(* PLC project PR_5by3CylModWoRdlck_PLC, SiemensToBackhoff Siemens TIA Portal to Beckhoff TwinCAT PLCopen Converter 2.0 *)
(* stored: creationDateTime 2026-09-28T12:19:39.070834, modificationDateTime 2026-09-28T12:19:39.070834 *)

FUNCTION_BLOCK PR_5by3CylModWoRdlck
VAR_INPUT
	iResetModule : BOOL;  // Reset if 1
	iResetFaults : BOOL;  // Reset Fault CMD
	iEnergizeAtPwrOn : BOOL;  // Energize Poweron Input
	iWorkCmd : BOOL;  // Cyl Work Postion CMD
	iHomeCmd : BOOL;  // Cyl Home Postion CMD
	iWorkSen : BOOL;  // Cyl Work Postion Input
	iHomeSen : BOOL;  // Cyl Home Postion Input
	iWorkCleartoMove : BOOL;  // connect work position interlock condition healthy
	iHomeCleartoMove : BOOL;  // connect home position interlock condition healthy
	iWorkPositionLeftOption : BOOL;  // It is the selection of the to keep work solenoid coil on after reaching work position
	iHomePositionLeftOption : BOOL;  // It is the selection of the to keep home solenoid coil on after reaching home position
	iTimeoutValue : TIME;  // Time Required E.g T#500MS,T#2S
	iWorkSensDebounceVal : TIME;  // Time Required E.g T#500MS,T#2S
	iHomeSensDebounceVal : TIME;  // Time Required E.g T#500MS,T#2S
END_VAR
VAR_OUTPUT
	qWorkSol : BOOL;  // Cyl Work Position Sol Output
	qHomeSol : BOOL;  // Cyl Home Position Sol Output
	qWorkOver : BOOL;  // 1 if Cyl at Work Position
	qHomeOver : BOOL;  // 1 if Cyl at Home Position
	qModError : BOOL;  // Module Error
	qErrBothSensorOn : BOOL;  // 1 If both WorkSen and HomeSen inputs are high at the same time.
	qErrHomeInterlock : BOOL;  // 1 If homeCleartoMove is low and home command is active.
	qErrHomeSenNotLeft : BOOL;  // 1 If home position sensor did not turn off within defined time
	qErrHomeTout : BOOL;  // 1 If cylinder did not reach home position within defined time
	qErrWorkInterlock : BOOL;  // 1 If WorkCleartoMove is low and work command is active.
	qErrWorkSenNotLeft : BOOL;  // 1 If work position sensor did not turn off within defined time
	qErrWorkTout : BOOL;  // 1 If cylinder did not reach work position within defined time
	qMsgWorkPosLost : BOOL;  // 1 If work position achieved and lost its position without home
	qMsgHomePosLost : BOOL;  // 1 If home position achieved and lost its position without work
	qMsgBothCmdOn : BOOL;  // 1 if Home & work position command on same time
END_VAR
VAR
	sFltRstPls : BOOL;  // Stat bit for positive edge of reset fault input
	sFltEdge : R_TRIG;  // Positive edge of fault reset input
	sWorkPosMemBit : BOOL;  // Stat bit for work position memory bit
	sHomePosMemBit : BOOL;  // Stat bit for Home position memory bit
	sModError : BOOL;  // Stat bit for Module error
	sWorkSensDebTime : TIME;  // Stat bit work sensor debounce time
	sHomeSensDebTime : TIME;  // Stat bit work sensor debounce time
	sTimeoutValue : TIME;  // Stat bit for time out value
	sElapsedTime : TIME;  // Stat bit for time elapsed
	sDlyWorkSensDeb : TON;  // On Delay for Work Sensor Debounce
	sDlyHomeSensDeb : TON;  // On Delay For Home Sensor Debounce
	sDlyTimeOut : TON;  // On Delay Time Out timer
	sWorkSol : BOOL;
	sErrWorkTout : BOOL;
	sHomeSol : BOOL;
	sErrHomeTout : BOOL;
	sErrBothSensorOn : BOOL;
	sErrWorkInterlock : BOOL;
	sErrHomeInterlock : BOOL;
	sErrWorkSenNotLeft : BOOL;
	sErrHomeSenNotLeft : BOOL;
	sMsgHomePosLost : BOOL;
	sMsgWorkPosLost : BOOL;
	sPosEdge : R_TRIG;
	sPosEdge1 : R_TRIG;
	sRegainWrkPos : BOOL;
	sRegainHomePos : BOOL;
	sBothCmdOn : BOOL;
	sWorkPositionLeft : BOOL;
	sHomePositionLeft : BOOL;
END_VAR
  VAR  (* added by the conversion: wires and edge detectors of the diagram *)
    _EQ31_ENO : BOOL;
    _EQ31_OUT : BOOL;
    _EQ47_ENO : BOOL;
    _EQ47_OUT : BOOL;
    _EQ63_ENO : BOOL;
    _EQ63_OUT : BOOL;
  END_VAR

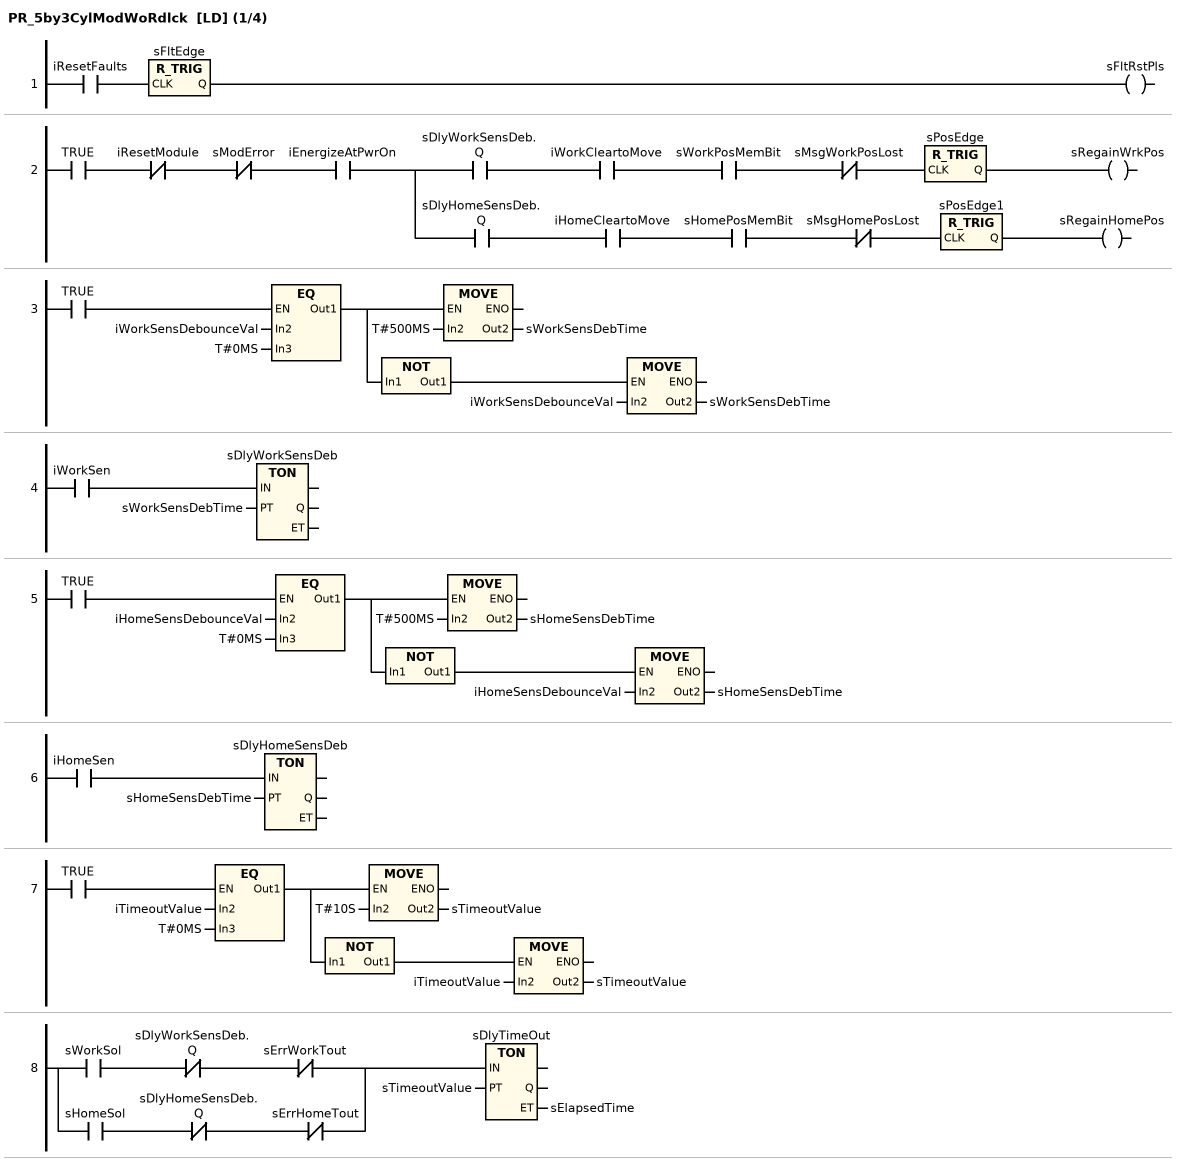
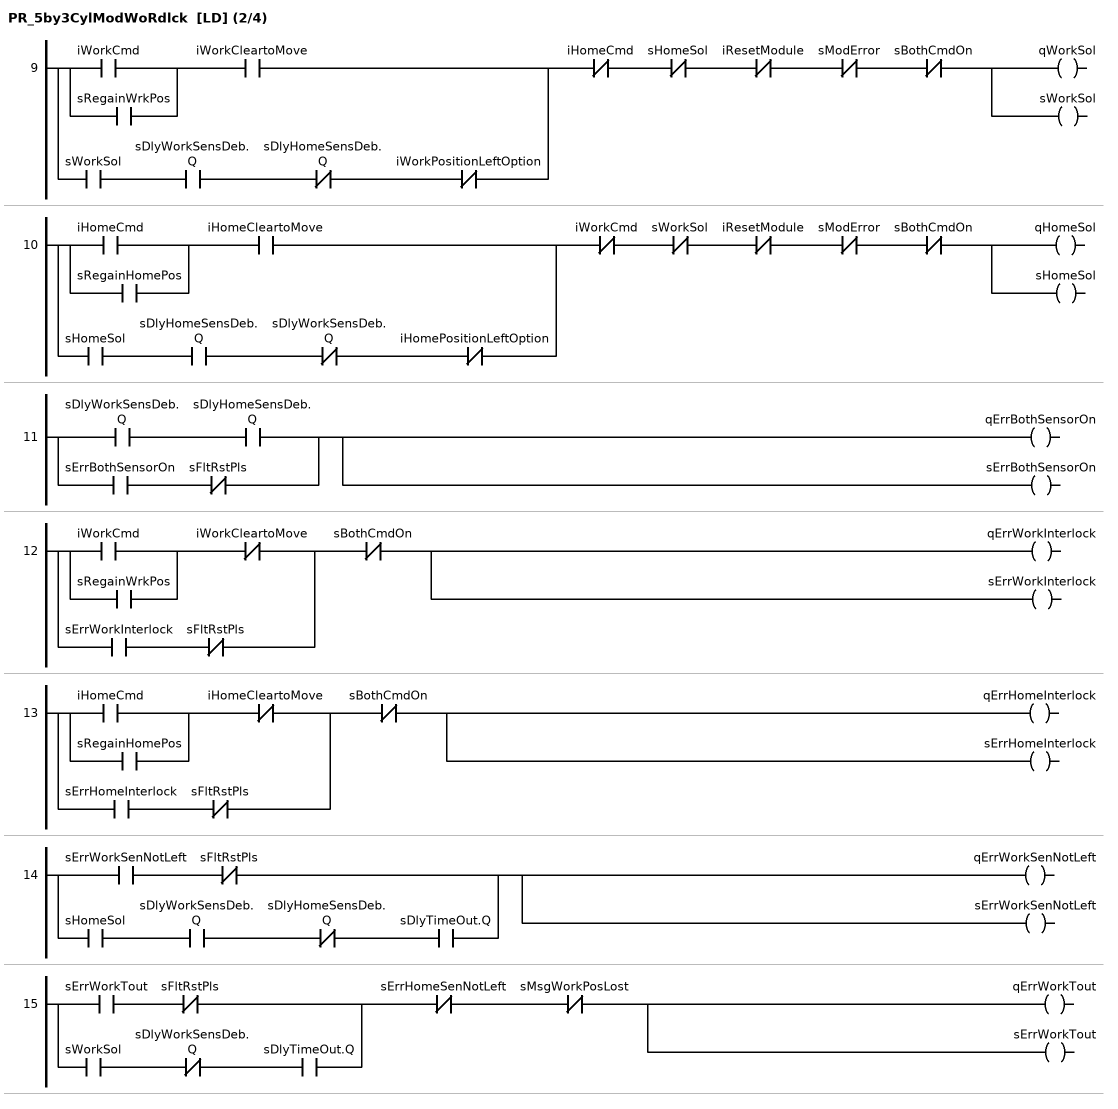
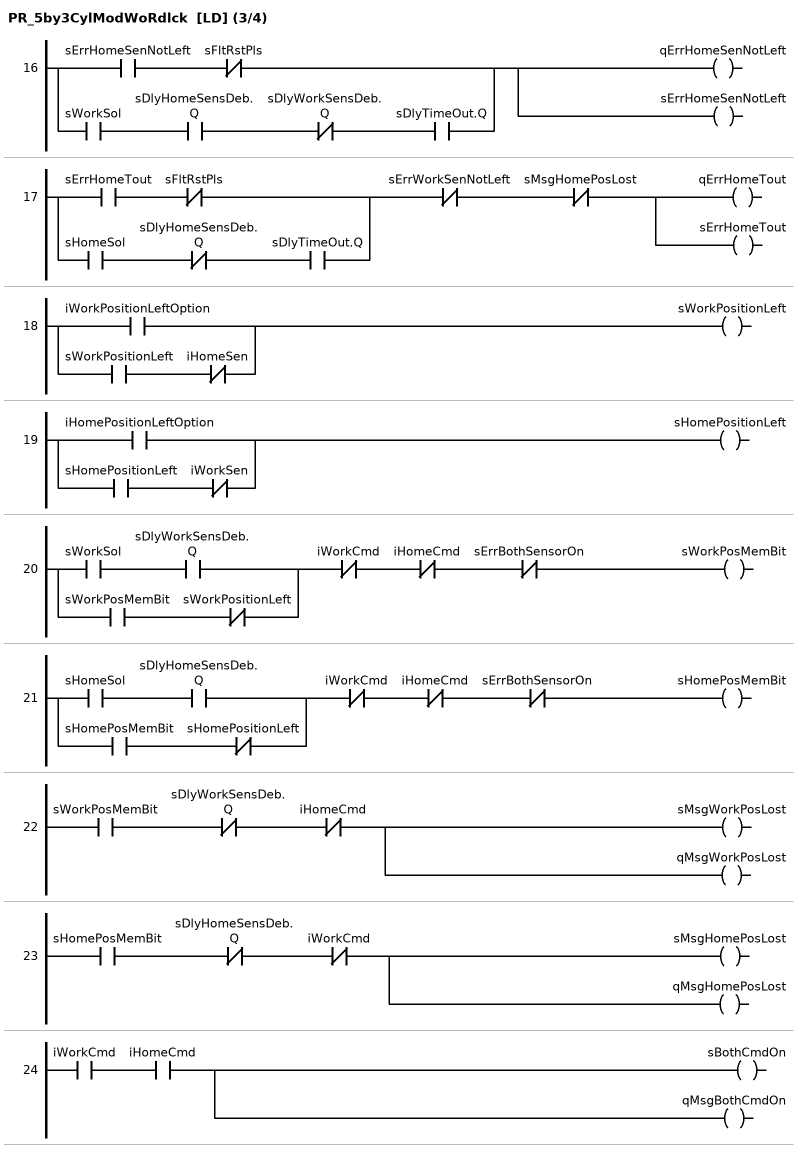
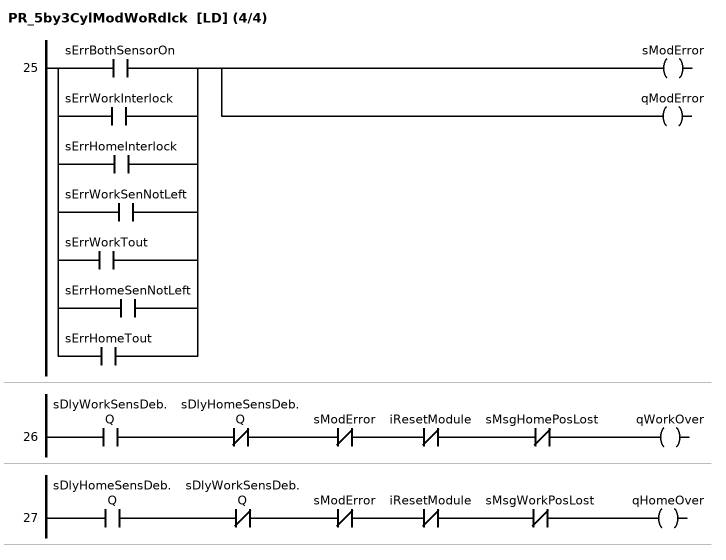
(* LD diagram, written out as Structured Text *)
(* ==============================================================================
 Company: Precision Automation & Robotics India Ltd. 
------------------------------------------------------------------------------
 Item Code:SM0101022005
 Author/Created by: Amiya Das
 Reviewed/Checked by: Atul Patwardhan
 First Release on: 20-01-2017
 Latest update on:27-01-2025 
------------------------------------------------------------------------------
 Tested with:Simulator
 Engineering/Editor: TIA Portal 15 & Higher
------------------------------------------------------------------------------
 Restrictions: No
 Dependencies/Requirements: NA
------------------------------------------------------------------------------
 Change Log:
 Ver.	Date                            Changed by                                  Details of changes
 0.2           20-01-2017                  Amiya Das      	              Second release version
 0.3           27-01-2025                 Sujeet Rote                                qMsgBothCmdOn message is added
 0.4           29-01-2025                  Sujeet Rote                                Work & home position left option bit
------------------------------------------------------------------------------
Functionality: This block is used to control a simple motion with one work 
position output, one home position  output, one work position sensor and one 
home position sensor.
Inputs
iResetModule	Bool
iResetFaults	Bool
iEnergizeAtPwrOn	Bool
iWorkCmd	Bool
iHomeCmd	Bool
iWorkSen	Bool
iHomeSen	Bool
iWorkCleartoMove	Bool
iHomeCleartoMove	Bool
iWorkPositionLeftOption	Bool
iHomePositionLeftOption	Bool
iTimeoutValue	Time
iWorkSensDebounceVal	Time
iHomeSensDebounceVal	Time

Outputs
qWorkSol	Bool
qHomeSol	Bool
qWorkOver	Bool
qHomeOver	Bool
qErrBothSensorOn	Bool
qErrHomeInterlock	Bool
qErrHomeSenNotLeft	Bool
qErrHomeTout	Bool
qErrWorkInterlock	Bool
qErrWorkSenNotLeft	Bool
qErrWorkTout	Bool
qMsgWorkPosLost	Bool
qMsgHomePosLost	Bool
qMsgBothCmdOn	Bool

In-outs
NIL
------------------------------------------------------------------------------
Errors reported:
1.qErrBothSensorOn: If both WorkSen and HomeSen inputs are high at the same time.          
2.qErrHomeInterlock: If homeCleartoMove is low and home command is active.
3.qErrHomeSenNotLeft: If home position sensor did not turn off within defined time 
4.qErrHomeTout: If cylinder did not reach home position within defined time 
5.qErrWorkInterlock: If WorkCleartoMove is low and work command is active. 
7.qErrWorkSenNotLeft: If work position sensor did not turn off within defined time 
8.qErrWorkTout: If cylinder did not reach work position within defined time 
9.qErrPipeSwaped: If Pipe or sensor swapped

Messages reported:
1.qMsgHomePosLost: If home position achieved and lost its position without work
2.qMsgWorkPosLost: If work position achieved and lost its position without home 
3.qMsgBothCmdOn :  Home & work position command on same time
============================================================================== *)

(* Fault Reset Pulse *)

sFltEdge(CLK := iResetFaults);
sFltRstPls := sFltEdge.Q;
(* Regain Position after power On logic *)

sPosEdge(CLK := TRUE AND NOT iResetModule AND NOT sModError AND iEnergizeAtPwrOn AND sDlyWorkSensDeb.Q AND iWorkCleartoMove AND sWorkPosMemBit AND NOT sMsgWorkPosLost);
sRegainWrkPos := sPosEdge.Q;
sPosEdge1(CLK := TRUE AND NOT iResetModule AND NOT sModError AND iEnergizeAtPwrOn AND sDlyHomeSensDeb.Q AND iHomeCleartoMove AND sHomePosMemBit AND NOT sMsgHomePosLost);
sRegainHomePos := sPosEdge1.Q;
(* Work sensor default debounce value *)

_EQ31_OUT := EQ(EN := TRUE, IN1 := iWorkSensDebounceVal, IN2 := T#0MS, ENO => _EQ31_ENO);
IF _EQ31_OUT THEN sWorkSensDebTime := T#500MS; END_IF;
IF NOT _EQ31_OUT THEN sWorkSensDebTime := iWorkSensDebounceVal; END_IF;
(* Work Sensor On Debounce Timer *)

sDlyWorkSensDeb(IN := iWorkSen, PT := sWorkSensDebTime);
(* Home sensor default debounce value *)

_EQ47_OUT := EQ(EN := TRUE, IN1 := iHomeSensDebounceVal, IN2 := T#0MS, ENO => _EQ47_ENO);
IF _EQ47_OUT THEN sHomeSensDebTime := T#500MS; END_IF;
IF NOT _EQ47_OUT THEN sHomeSensDebTime := iHomeSensDebounceVal; END_IF;
(* Home Sensor On Debounce Timer *)

sDlyHomeSensDeb(IN := iHomeSen, PT := sHomeSensDebTime);
(* Timeout Value *)

_EQ63_OUT := EQ(EN := TRUE, IN1 := iTimeoutValue, IN2 := T#0MS, ENO => _EQ63_ENO);
IF _EQ63_OUT THEN sTimeoutValue := T#10S; END_IF;
IF NOT _EQ63_OUT THEN sTimeoutValue := iTimeoutValue; END_IF;
(* Sensor timeout Timer *)

sDlyTimeOut(IN := sWorkSol AND NOT sDlyWorkSensDeb.Q AND NOT sErrWorkTout OR sHomeSol AND NOT sDlyHomeSensDeb.Q AND NOT sErrHomeTout, PT := sTimeoutValue, ET => sElapsedTime);
(* Cylinder Work Sol *)

qWorkSol := ((iWorkCmd OR sRegainWrkPos) AND iWorkCleartoMove OR sWorkSol AND sDlyWorkSensDeb.Q AND NOT sDlyHomeSensDeb.Q AND NOT iWorkPositionLeftOption) AND NOT iHomeCmd AND NOT sHomeSol AND NOT iResetModule AND NOT sModError AND NOT sBothCmdOn;
sWorkSol := ((iWorkCmd OR sRegainWrkPos) AND iWorkCleartoMove OR sWorkSol AND sDlyWorkSensDeb.Q AND NOT sDlyHomeSensDeb.Q AND NOT iWorkPositionLeftOption) AND NOT iHomeCmd AND NOT sHomeSol AND NOT iResetModule AND NOT sModError AND NOT sBothCmdOn;
(* Cylinder Home Sol *)

qHomeSol := ((iHomeCmd OR sRegainHomePos) AND iHomeCleartoMove OR sHomeSol AND sDlyHomeSensDeb.Q AND NOT sDlyWorkSensDeb.Q AND NOT iHomePositionLeftOption) AND NOT iWorkCmd AND NOT sWorkSol AND NOT iResetModule AND NOT sModError AND NOT sBothCmdOn;
sHomeSol := ((iHomeCmd OR sRegainHomePos) AND iHomeCleartoMove OR sHomeSol AND sDlyHomeSensDeb.Q AND NOT sDlyWorkSensDeb.Q AND NOT iHomePositionLeftOption) AND NOT iWorkCmd AND NOT sWorkSol AND NOT iResetModule AND NOT sModError AND NOT sBothCmdOn;
(* Both Sensor On Error *)

qErrBothSensorOn := sDlyWorkSensDeb.Q AND sDlyHomeSensDeb.Q OR sErrBothSensorOn AND NOT sFltRstPls;
sErrBothSensorOn := sDlyWorkSensDeb.Q AND sDlyHomeSensDeb.Q OR sErrBothSensorOn AND NOT sFltRstPls;
(* Work Interlock Error *)

qErrWorkInterlock := ((iWorkCmd OR sRegainWrkPos) AND NOT iWorkCleartoMove OR sErrWorkInterlock AND NOT sFltRstPls) AND NOT sBothCmdOn;
sErrWorkInterlock := ((iWorkCmd OR sRegainWrkPos) AND NOT iWorkCleartoMove OR sErrWorkInterlock AND NOT sFltRstPls) AND NOT sBothCmdOn;
(* Home Interlock Error pending *)

qErrHomeInterlock := ((iHomeCmd OR sRegainHomePos) AND NOT iHomeCleartoMove OR sErrHomeInterlock AND NOT sFltRstPls) AND NOT sBothCmdOn;
sErrHomeInterlock := ((iHomeCmd OR sRegainHomePos) AND NOT iHomeCleartoMove OR sErrHomeInterlock AND NOT sFltRstPls) AND NOT sBothCmdOn;
(* Work Sensor Not Left Error  pending *)

qErrWorkSenNotLeft := sHomeSol AND sDlyWorkSensDeb.Q AND NOT sDlyHomeSensDeb.Q AND sDlyTimeOut.Q OR sErrWorkSenNotLeft AND NOT sFltRstPls;
sErrWorkSenNotLeft := sHomeSol AND sDlyWorkSensDeb.Q AND NOT sDlyHomeSensDeb.Q AND sDlyTimeOut.Q OR sErrWorkSenNotLeft AND NOT sFltRstPls;
(* Work Timeout Error *)

qErrWorkTout := (sWorkSol AND NOT sDlyWorkSensDeb.Q AND sDlyTimeOut.Q OR sErrWorkTout AND NOT sFltRstPls) AND NOT sErrHomeSenNotLeft AND NOT sMsgWorkPosLost;
sErrWorkTout := (sWorkSol AND NOT sDlyWorkSensDeb.Q AND sDlyTimeOut.Q OR sErrWorkTout AND NOT sFltRstPls) AND NOT sErrHomeSenNotLeft AND NOT sMsgWorkPosLost;
(* Home Sensor Not Left Error *)

qErrHomeSenNotLeft := sWorkSol AND sDlyHomeSensDeb.Q AND NOT sDlyWorkSensDeb.Q AND sDlyTimeOut.Q OR sErrHomeSenNotLeft AND NOT sFltRstPls;
sErrHomeSenNotLeft := sWorkSol AND sDlyHomeSensDeb.Q AND NOT sDlyWorkSensDeb.Q AND sDlyTimeOut.Q OR sErrHomeSenNotLeft AND NOT sFltRstPls;
(* Home Timeout Error *)

qErrHomeTout := (sHomeSol AND NOT sDlyHomeSensDeb.Q AND sDlyTimeOut.Q OR sErrHomeTout AND NOT sFltRstPls) AND NOT sErrWorkSenNotLeft AND NOT sMsgHomePosLost;
sErrHomeTout := (sHomeSol AND NOT sDlyHomeSensDeb.Q AND sDlyTimeOut.Q OR sErrHomeTout AND NOT sFltRstPls) AND NOT sErrWorkSenNotLeft AND NOT sMsgHomePosLost;
(* Work Position Left option bit Logic *)

sWorkPositionLeft := iWorkPositionLeftOption OR sWorkPositionLeft AND NOT iHomeSen;
(* Home Position Left option bit Logic *)

sHomePositionLeft := iHomePositionLeftOption OR sHomePositionLeft AND NOT iWorkSen;
(* Work Position Memory Bit *)

sWorkPosMemBit := (sWorkSol AND sDlyWorkSensDeb.Q OR sWorkPosMemBit AND NOT sWorkPositionLeft) AND NOT iWorkCmd AND NOT iHomeCmd AND NOT sErrBothSensorOn;
(* Home Position Memory Bit *)

sHomePosMemBit := (sHomeSol AND sDlyHomeSensDeb.Q OR sHomePosMemBit AND NOT sHomePositionLeft) AND NOT iWorkCmd AND NOT iHomeCmd AND NOT sErrBothSensorOn;
(* Msg:-Work Position Lost *)

sMsgWorkPosLost := sWorkPosMemBit AND NOT sDlyWorkSensDeb.Q AND NOT iHomeCmd;
qMsgWorkPosLost := sWorkPosMemBit AND NOT sDlyWorkSensDeb.Q AND NOT iHomeCmd;
(* Msg:- Home Position Lost *)

sMsgHomePosLost := sHomePosMemBit AND NOT sDlyHomeSensDeb.Q AND NOT iWorkCmd;
qMsgHomePosLost := sHomePosMemBit AND NOT sDlyHomeSensDeb.Q AND NOT iWorkCmd;
(* Msg:- Both command On *)

sBothCmdOn := iWorkCmd AND iHomeCmd;
qMsgBothCmdOn := iWorkCmd AND iHomeCmd;
(* Module Error *)

sModError := sErrBothSensorOn OR sErrWorkInterlock OR sErrHomeInterlock OR sErrWorkSenNotLeft OR sErrWorkTout OR sErrHomeSenNotLeft OR sErrHomeTout;
qModError := sErrBothSensorOn OR sErrWorkInterlock OR sErrHomeInterlock OR sErrWorkSenNotLeft OR sErrWorkTout OR sErrHomeSenNotLeft OR sErrHomeTout;
(* Work Over *)

qWorkOver := sDlyWorkSensDeb.Q AND NOT sDlyHomeSensDeb.Q AND NOT sModError AND NOT iResetModule AND NOT sMsgHomePosLost;
(* Home Over *)

qHomeOver := sDlyHomeSensDeb.Q AND NOT sDlyWorkSensDeb.Q AND NOT sModError AND NOT iResetModule AND NOT sMsgWorkPosLost;
END_FUNCTION_BLOCK
